// TIA Portal V17 export
FUNCTION "FC_T05_Boites" : Void   // FC105, LAD
{ S7_Optimized_Access := 'TRUE' }
// stored: SetENOAutomatically false
   VAR_INPUT
      Valeur_A : Int;
      Valeur_B : Int;
   END_VAR
   VAR_OUTPUT
      Copie : Int;
      Somme : Int;
      Superieur_Egal : Bool;
      Egal : Bool;
   END_VAR
BEGIN

REGION Network 1: MOVE
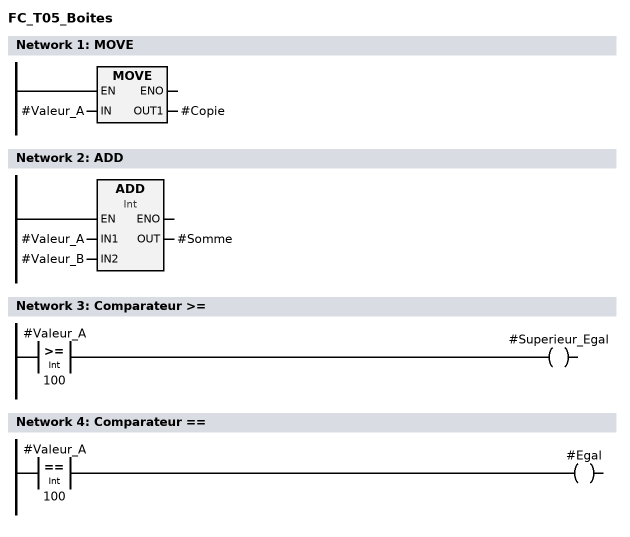
   RUNG wire#powerrail
      Move(in := #Valeur_A, out1 => #Copie)
   END_RUNG
   // the same network as SCL:
   #Copie := #Valeur_A;
END_REGION

REGION Network 2: ADD
   RUNG wire#powerrail
      { S7_Templates := "SrcType := Int" } Add(in1 := #Valeur_A, in2 := #Valeur_B, out => #Somme)
   END_RUNG
   // the same network as SCL:
   #Somme := #Valeur_A + #Valeur_B;
END_REGION

REGION Network 3: Comparateur >=
   RUNG wire#powerrail
      { S7_Templates := "SrcType := Int" } GE_Contact(in1 := #Valeur_A, in2 := 100)
      Coil( #Superieur_Egal )
   END_RUNG
   // the same network as SCL:
   #Superieur_Egal := #Valeur_A >= 100;
END_REGION

REGION Network 4: Comparateur ==
   RUNG wire#powerrail
      { S7_Templates := "SrcType := Int" } EQ_Contact(in1 := #Valeur_A, in2 := 100)
      Coil( #Egal )
   END_RUNG
   // the same network as SCL:
   #Egal := #Valeur_A = 100;
END_REGION
END_FUNCTION
